// TIA Portal V21 export
// export: Created 2026-11-21T12:56:43.283546Z, ExportSetting WithDefaults, DisplayName Totally Integrated Automation Portal, DisplayVersion V21, DisplayName STEP 7 Professional, DisplayVersion V21, DisplayName STEP 7 Safety, DisplayVersion V21, DisplayName Tech WebApplication, DisplayVersion V21, DisplayName WinCC Basic/Comfort/Advanced, DisplayVersion V21, DisplayName WinCC Unified, DisplayVersion V21
VAR_GLOBAL   // PLC tag table "IO"
   Start_Partner AT %I0.0 : Bool;   // An input of the partner
   Lamp_Partner AT %Q0.0 : Bool;   // First output of Outputs_P
END_VAR
